            mdesc mMdesc
            num nActionIndex
            num nDelay = 0.5
            num nMoveType = 7
            num nPercentage
            num nSigValue
        pointRx pPointRx[2]
        string sID
      [5]
        bool bMarked
        jointRx jJointRx
        pointRx pInter
        paraItem pParaItem
          [0]
            bool bSafePoint
            ifItem iIfItem
              [0]
                bool bANDOR[2]
                num nSigIndex[3]
                num nSigType[3]
                num nValue[3]
            mdesc mMdesc
            num nActionIndex = 40
            num nDelay
            num nMoveType = 4
            num nPercentage
            num nSigValue
        pointRx pPointRx[2]
        string sID
    string sID
  [Y006]
    num nFrameIndex
    num nMoveID
    num nToolIndex
    pointItem pPointItem[6]
      [0]
        bool bMarked
        jointRx jJointRx
        pointRx pInter
        paraItem pParaItem
          [0]
            bool bSafePoint
            ifItem iIfItem
              [0]
                bool bANDOR[2]
                num nSigIndex[3]
                num nSigType[3]
                num nValue[3]
            mdesc mMdesc
            num nActionIndex = 40
            num nDelay
            num nMoveType = 4
            num nPercentage
            num nSigValue = 1
        pointRx pPointRx[2]
        string sID
      [1]
        bool bMarked
        jointRx jJointRx
        pointRx pInter
        paraItem pParaItem
          [0]
            bool bSafePoint
            ifItem iIfItem
              [0]
                bool bANDOR[2]
                num nSigIndex[3]
                num nSigType[3]
                num nValue[3]
            mdesc mMdesc
            num nActionIndex = 5
            num nDelay
            num nMoveType = 6
            num nPercentage
            num nSigValue = 6
        pointRx pPointRx[2]
        string sID
      [2]
        bool bMarked
        jointRx jJointRx
        pointRx pInter
        paraItem pParaItem
          [0]
            bool bSafePoint
            ifItem iIfItem
              [0]
                bool bANDOR[2]
                num nSigIndex[3]
                num nSigType[3]
                num nValue[3]
            mdesc mMdesc
            num nActionIndex
            num nDelay = 0.5
            num nMoveType = 7
            num nPercentage
            num nSigValue
        pointRx pPointRx[2]
        string sID
      [3]
        bool bMarked
        jointRx jJointRx
        pointRx pInter
        paraItem pParaItem
          [0]
            bool bSafePoint
            ifItem iIfItem
              [0]
                bool bANDOR[2]
                num nSigIndex[3]
                num nSigType[3]
                num nValue[3]
            mdesc mMdesc
            num nActionIndex = 40
            num nDelay = 0.5
            num nMoveType = 3
            num nPercentage
            num nSigValue = 1
        pointRx pPointRx[2]
        string sID
      [4]
        bool bMarked
        jointRx jJointRx
        pointRx pInter
        paraItem pParaItem
          [0]
            bool bSafePoint
            ifItem iIfItem
              [0]
                bool bANDOR[2]
                num nSigIndex[3]
                num nSigType[3]
                num nValue[3]
            mdesc mMdesc
            num nActionIndex
            num nDelay = 0.5
            num nMoveType = 7
            num nPercentage
            num nSigValue
        pointRx pPointRx[2]
        string sID
      [5]
        bool bMarked
        jointRx jJointRx
        pointRx pInter
        paraItem pParaItem
          [0]
            bool bSafePoint
            ifItem iIfItem
              [0]
                bool bANDOR[2]
                num nSigIndex[3]
                num nSigType[3]
                num nValue[3]
            mdesc mMdesc
            num nActionIndex = 40
            num nDelay
            num nMoveType = 4
            num nPercentage
            num nSigValue
        pointRx pPointRx[2]
        string sID
    string sID
  [Y007]
    num nFrameIndex
    num nMoveID
    num nToolIndex
    pointItem pPointItem[6]
      [0]
        bool bMarked
        jointRx jJointRx
        pointRx pInter
        paraItem pParaItem
          [0]
            bool bSafePoint
            ifItem iIfItem
              [0]
                bool bANDOR[2]
                num nSigIndex[3]
                num nSigType[3]
                num nValue[3]
            mdesc mMdesc
            num nActionIndex = 40
            num nDelay
            num nMoveType = 4
            num nPercentage
            num nSigValue = 1
        pointRx pPointRx[2]
        string sID
      [1]
        bool bMarked
        jointRx jJointRx
        pointRx pInter
        paraItem pParaItem
          [0]
            bool bSafePoint
            ifItem iIfItem
              [0]
                bool bANDOR[2]
                num nSigIndex[3]
                num nSigType[3]
                num nValue[3]
            mdesc mMdesc
            num nActionIndex = 5
            num nDelay
            num nMoveType = 6
            num nPercentage
            num nSigValue = 7
        pointRx pPointRx[2]
        string sID
      [2]
        bool bMarked
        jointRx jJointRx
        pointRx pInter
        paraItem pParaItem
          [0]
            bool bSafePoint
            ifItem iIfItem
              [0]
                bool bANDOR[2]
                num nSigIndex[3]
                num nSigType[3]
                num nValue[3]
            mdesc mMdesc
            num nActionIndex
            num nDelay = 0.5
            num nMoveType = 7
            num nPercentage
            num nSigValue
        pointRx pPointRx[2]
        string sID
      [3]
        bool bMarked
        jointRx jJointRx
        pointRx pInter
        paraItem pParaItem
          [0]
            bool bSafePoint
            ifItem iIfItem
              [0]
                bool bANDOR[2]
                num nSigIndex[3]
                num nSigType[3]
                num nValue[3]
            mdesc mMdesc
            num nActionIndex = 40
            num nDelay = 0.5
            num nMoveType = 3
            num nPercentage
            num nSigValue = 1
        pointRx pPointRx[2]
        string sID
      [4]
        bool bMarked
        jointRx jJointRx
        pointRx pInter
        paraItem pParaItem
          [0]
            bool bSafePoint
            ifItem iIfItem
              [0]
                bool bANDOR[2]
                num nSigIndex[3]
                num nSigType[3]
                num nValue[3]
            mdesc mMdesc
            num nActionIndex
            num nDelay = 0.5
            num nMoveType = 7
            num nPercentage
            num nSigValue
        pointRx pPointRx[2]
        string sID
      [5]
        bool bMarked
        jointRx jJointRx
        pointRx pInter
        paraItem pParaItem
          [0]
            bool bSafePoint
            ifItem iIfItem
              [0]
                bool bANDOR[2]
                num nSigIndex[3]
                num nSigType[3]
                num nValue[3]
            mdesc mMdesc
            num nActionIndex = 40
            num nDelay
            num nMoveType = 4
            num nPercentage
            num nSigValue
        pointRx pPointRx[2]
        string sID
    string sID
  [Y008]
    num nFrameIndex
    num nMoveID
    num nToolIndex
    pointItem pPointItem[6]
      [0]
        bool bMarked
        jointRx jJointRx
        pointRx pInter
        paraItem pParaItem
          [0]
            bool bSafePoint
            ifItem iIfItem
              [0]
                bool bANDOR[2]
                num nSigIndex[3]
                num nSigType[3]
                num nValue[3]
            mdesc mMdesc
            num nActionIndex = 40
            num nDelay
            num nMoveType = 4
            num nPercentage
            num nSigValue = 1
        pointRx pPointRx[2]
        string sID
      [1]
        bool bMarked
        jointRx jJointRx
        pointRx pInter
        paraItem pParaItem
          [0]
            bool bSafePoint
            ifItem iIfItem
              [0]
                bool bANDOR[2]
                num nSigIndex[3]
                num nSigType[3]
                num nValue[3]
            mdesc mMdesc
            num nActionIndex = 5
            num nDelay
            num nMoveType = 6
            num nPercentage
            num nSigValue = 8
        pointRx pPointRx[2]
        string sID
      [2]
        bool bMarked
        jointRx jJointRx
        pointRx pInter
        paraItem pParaItem
          [0]
            bool bSafePoint
            ifItem iIfItem
              [0]
                bool bANDOR[2]
                num nSigIndex[3]
                num nSigType[3]
                num nValue[3]
            mdesc mMdesc
            num nActionIndex
            num nDelay = 0.5
            num nMoveType = 7
            num nPercentage
            num nSigValue
        pointRx pPointRx[2]
        string sID
      [3]
        bool bMarked
        jointRx jJointRx
        pointRx pInter
        paraItem pParaItem
          [0]
            bool bSafePoint
            ifItem iIfItem
              [0]
                bool bANDOR[2]
                num nSigIndex[3]
                num nSigType[3]
                num nValue[3]
            mdesc mMdesc
            num nActionIndex = 40
            num nDelay = 0.5
            num nMoveType = 3
            num nPercentage
            num nSigValue = 1
        pointRx pPointRx[2]
        string sID
      [4]
        bool bMarked
        jointRx jJointRx
        pointRx pInter
        paraItem pParaItem
          [0]
            bool bSafePoint
            ifItem iIfItem
              [0]
                bool bANDOR[2]
                num nSigIndex[3]
                num nSigType[3]
                num nValue[3]
            mdesc mMdesc
            num nActionIndex
            num nDelay = 0.5
            num nMoveType = 7
            num nPercentage
            num nSigValue
        pointRx pPointRx[2]
        string sID
      [5]
        bool bMarked
        jointRx jJointRx
        pointRx pInter
        paraItem pParaItem
          [0]
            bool bSafePoint
            ifItem iIfItem
              [0]
                bool bANDOR[2]
                num nSigIndex[3]
                num nSigType[3]
                num nValue[3]
            mdesc mMdesc
            num nActionIndex = 40
            num nDelay
            num nMoveType = 4
            num nPercentage
            num nSigValue
        pointRx pPointRx[2]
        string sID
    string sID
  [complete]
    num nFrameIndex
    num nMoveID
    num nToolIndex
    pointItem pPointItem[3]
      [0]
        bool bMarked
        jointRx jJointRx
        pointRx pInter
        paraItem pParaItem
          [0]
            bool bSafePoint
            ifItem iIfItem
              [0]
                bool bANDOR[2]
                num nSigIndex[3]
                num nSigType[3]
                num nValue[3]
            mdesc mMdesc
            num nActionIndex = 50
            num nDelay
            num nMoveType = 4
            num nPercentage
            num nSigValue = 1
        pointRx pPointRx[2]
        string sID
      [1]
        bool bMarked
        jointRx jJointRx
        pointRx pInter
        paraItem pParaItem
          [0]
            bool bSafePoint
            ifItem iIfItem
              [0]
                bool bANDOR[2]
                num nSigIndex[3]
                num nSigType[3]
                num nValue[3]
            mdesc mMdesc
            num nActionIndex = 50
            num nDelay = 3
            num nMoveType = 7
            num nPercentage
            num nSigValue = 1
        pointRx pPointRx[2]
        string sID
      [2]
        bool bMarked
        jointRx jJointRx
        pointRx pInter
        paraItem pParaItem
          [0]
            bool bSafePoint
            ifItem iIfItem
              [0]
                bool bANDOR[2]
                num nSigIndex[3]
                num nSigType[3]
                num nValue[3]
            mdesc mMdesc
            num nActionIndex = 50
            num nDelay = 3
            num nMoveType = 4
            num nPercentage
            num nSigValue
        pointRx pPointRx[2]
        string sID
    string sID
  [gggg]
    num nFrameIndex
    num nMoveID
    num nToolIndex
    pointItem pPointItem
      [0]
        bool bMarked
        jointRx jJointRx
        pointRx pInter
        paraItem pParaItem
          [0]
            bool bSafePoint
            ifItem iIfItem
              [0]
                bool bANDOR[2]
                num nSigIndex[3]
                num nSigType[3]
                num nValue[3]
            mdesc mMdesc
            num nActionIndex
            num nDelay
            num nMoveType
            num nPercentage
            num nSigValue
        pointRx pPointRx[2]
        string sID
    string sID
  [init]
    num nFrameIndex
    num nMoveID
    num nToolIndex
    pointItem pPointItem[14]
      [0]
        bool bMarked
        jointRx jJointRx
        pointRx pInter
        paraItem pParaItem
          [0]
            bool bSafePoint
            ifItem iIfItem
              [0]
                bool bANDOR[2]
                num nSigIndex[3]
                num nSigType[3]
                num nValue[3]
            mdesc mMdesc
            num nActionIndex
            num nDelay
            num nMoveType = 6
            num nPercentage
            num nSigValue
        pointRx pPointRx[2]
        string sID
      [1]
        bool bMarked
        jointRx jJointRx
        pointRx pInter
        paraItem pParaItem
          [0]
            bool bSafePoint
            ifItem iIfItem
              [0]
                bool bANDOR[2]
                num nSigIndex[3]
                num nSigType[3]
                num nValue[3]
            mdesc mMdesc
            num nActionIndex = 3
            num nDelay
            num nMoveType = 6
            num nPercentage
            num nSigValue
        pointRx pPointRx[2]
        string sID
      [2]
        bool bMarked
        jointRx jJointRx
        pointRx pInter
        paraItem pParaItem
          [0]
            bool bSafePoint
            ifItem iIfItem
              [0]
                bool bANDOR[2]
                num nSigIndex[3]
                num nSigType[3]
                num nValue[3]
            mdesc mMdesc
            num nActionIndex = 2
            num nDelay
            num nMoveType = 6
            num nPercentage
            num nSigValue
        pointRx pPointRx[2]
        string sID
      [3]
        bool bMarked
        jointRx jJointRx
        pointRx pInter
        paraItem pParaItem
          [0]
            bool bSafePoint
            ifItem iIfItem
              [0]
                bool bANDOR[2]
                num nSigIndex[3]
                num nSigType[3]
                num nValue[3]
            mdesc mMdesc
            num nActionIndex = 1
            num nDelay
            num nMoveType = 6
            num nPercentage
            num nSigValue
        pointRx pPointRx[2]
        string sID
      [4]
        bool bMarked
        jointRx jJointRx
        pointRx pInter
        paraItem pParaItem
          [0]
            bool bSafePoint
            ifItem iIfItem
              [0]
                bool bANDOR[2]
                num nSigIndex[3]
                num nSigType[3]
                num nValue[3]
            mdesc mMdesc
            num nActionIndex = 4
            num nDelay
            num nMoveType = 6
            num nPercentage
            num nSigValue
        pointRx pPointRx[2]
        string sID
      [5]
        bool bMarked
        jointRx jJointRx
        pointRx pInter
        paraItem pParaItem
          [0]
            bool bSafePoint
            ifItem iIfItem
              [0]
                bool bANDOR[2]
                num nSigIndex[3]
                num nSigType[3]
                num nValue[3]
            mdesc mMdesc
            num nActionIndex = 5
            num nDelay
            num nMoveType = 6
            num nPercentage
            num nSigValue
        pointRx pPointRx[2]
        string sID
      [6]
        bool bMarked
        jointRx jJointRx
        pointRx pInter
        paraItem pParaItem
          [0]
            bool bSafePoint
            ifItem iIfItem
              [0]
                bool bANDOR[2]
                num nSigIndex[3]
                num nSigType[3]
                num nValue[3]
            mdesc mMdesc
            num nActionIndex = 50
            num nDelay
            num nMoveType = 4
            num nPercentage
            num nSigValue
        pointRx pPointRx[2]
        string sID
      [7]
        bool bMarked
        jointRx jJointRx
        pointRx pInter
        paraItem pParaItem
          [0]
            bool bSafePoint
            ifItem iIfItem
              [0]
                bool bANDOR[2]
                num nSigIndex[3]
                num nSigType[3]
                num nValue[3]
            mdesc mMdesc
            num nActionIndex = 40
            num nDelay
            num nMoveType = 4
            num nPercentage
            num nSigValue
        pointRx pPointRx[2]
        string sID
      [8]
        bool bMarked
        jointRx jJointRx
        pointRx pInter
        paraItem pParaItem
          [0]
            bool bSafePoint
            ifItem iIfItem
              [0]
                bool bANDOR[2]
                num nSigIndex[3]
                num nSigType[3]
                num nValue[3]
            mdesc mMdesc
            num nActionIndex = 41
            num nDelay
            num nMoveType = 4
            num nPercentage
            num nSigValue
        pointRx pPointRx[2]
        string sID
      [9]
        bool bMarked
        jointRx jJointRx
        pointRx pInter
        paraItem pParaItem
          [0]
            bool bSafePoint
            ifItem iIfItem
              [0]
                bool bANDOR[2]
                num nSigIndex[3]
                num nSigType[3]
                num nValue[3]
            mdesc mMdesc
            num nActionIndex = 42
            num nDelay
            num nMoveType = 4
            num nPercentage
            num nSigValue
        pointRx pPointRx[2]
        string sID
      [10]
        bool bMarked
        jointRx jJointRx
        pointRx pInter
        paraItem pParaItem
          [0]
            bool bSafePoint
            ifItem iIfItem
              [0]
                bool bANDOR[2]
                num nSigIndex[3]
                num nSigType[3]
                num nValue[3]
            mdesc mMdesc
            num nActionIndex = 43
            num nDelay
            num nMoveType = 4
            num nPercentage
            num nSigValue
        pointRx pPointRx[2]
        string sID
      [11]
        bool bMarked
        jointRx jJointRx
        pointRx pInter
        paraItem pParaItem
          [0]
            bool bSafePoint
            ifItem iIfItem
              [0]
                bool bANDOR[2]
                num nSigIndex[3]
                num nSigType[3]
                num nValue[3]
            mdesc mMdesc
            num nActionIndex = 44
            num nDelay
            num nMoveType = 4
            num nPercentage
            num nSigValue
        pointRx pPointRx[2]
        string sID
      [12]
        bool bMarked
        jointRx jJointRx
        pointRx pInter
        paraItem pParaItem
          [0]
            bool bSafePoint
            ifItem iIfItem
              [0]
                bool bANDOR[2]
                num nSigIndex[3]
                num nSigType[3]
                num nValue[3]
            mdesc mMdesc
            num nActionIndex = 47
            num nDelay
            num nMoveType = 4
            num nPercentage
            num nSigValue
        pointRx pPointRx[2]
        string sID
      [13]
        bool bMarked
        jointRx jJointRx
        pointRx pInter
        paraItem pParaItem
          [0]
            bool bSafePoint
            ifItem iIfItem
              [0]
                bool bANDOR[2]
                num nSigIndex[3]
                num nSigType[3]
                num nValue[3]
            mdesc mMdesc
            num nActionIndex = 48
            num nDelay
            num nMoveType = 4
            num nPercentage
            num nSigValue
        pointRx pPointRx[2]
        string sID
    string sID
  [p001]
    num nFrameIndex
    num nMoveID
    num nToolIndex
    pointItem pPointItem[109]
      [0]
        bool bMarked
        jointRx jJointRx = {j1=14.463054, j2=126.686617, j3=-94.408556, j4=-18.307578, j5=-113.737208, j6=85.971215}
        pointRx pInter
        paraItem pParaItem
          [0]
            bool bSafePoint
            ifItem iIfItem
              [0]
                bool bANDOR[2]
                num nSigIndex[3]
                num nSigType[3]
                num nValue[3]
            mdesc mMdesc
            num nActionIndex = 41
            num nDelay = 1
            num nMoveType = 7
            num nPercentage
            num nSigValue
        pointRx pPointRx[2] = {x=278.890712, y=136.745171, z=230.948915, rx=84.337923, ry=-1.664851, rz=172.690172, shoulder=lefty, elbow=enegative, wrist=wnegative}
        string sID
      [1]
        bool bMarked
        jointRx jJointRx = {j1=14.463054, j2=126.686617, j3=-94.408556, j4=-18.307578, j5=-113.737208, j6=85.971215}
        pointRx pInter
        paraItem pParaItem
          [0]
            bool bSafePoint
            ifItem iIfItem
              [0]
                bool bANDOR[2]
                num nSigIndex[3]
                num nSigType[3]
                num nValue[3]
            mdesc mMdesc
            num nActionIndex = 71
            num nDelay = 1
            num nMoveType = 4
            num nPercentage
            num nSigValue
        pointRx pPointRx[2] = {x=278.890712, y=136.745171, z=230.948915, rx=84.337923, ry=-1.664851, rz=172.690172, shoulder=lefty, elbow=enegative, wrist=wnegative}
        string sID
      [2]
        bool bMarked
        jointRx jJointRx = {j1=14.463054, j2=126.686617, j3=-94.408556, j4=-18.307578, j5=-113.737208, j6=85.971215}
        pointRx pInter
        paraItem pParaItem
          [0]
            bool bSafePoint
            ifItem iIfItem
              [0]
                bool bANDOR[2]
                num nSigIndex[3]
                num nSigType[3]
                num nValue[3]
            mdesc mMdesc
            num nActionIndex = 70
            num nDelay = 1
            num nMoveType = 4
            num nPercentage
            num nSigValue = 1
        pointRx pPointRx[2] = {x=278.890712, y=136.745171, z=230.948915, rx=84.337923, ry=-1.664851, rz=172.690172, shoulder=lefty, elbow=enegative, wrist=wnegative}
        string sID
      [3]
        bool bMarked
        jointRx jJointRx = {j1=14.463054, j2=126.686617, j3=-94.408556, j4=-18.307578, j5=-113.737208, j6=85.971215}
        pointRx pInter
        paraItem pParaItem
          [0]
            bool bSafePoint
            ifItem iIfItem
              [0]
                bool bANDOR[2]
                num nSigIndex[3]
                num nSigType[3]
                num nValue[3]
            mdesc mMdesc
            num nActionIndex = 70
            num nDelay = 1
            num nMoveType = 3
            num nPercentage
            num nSigValue = 1
        pointRx pPointRx[2] = {x=278.890712, y=136.745171, z=230.948915, rx=84.337923, ry=-1.664851, rz=172.690172, shoulder=lefty, elbow=enegative, wrist=wnegative}
        string sID
      [4]
        bool bMarked
        jointRx jJointRx = {j1=-0.746077, j2=38.654193, j3=103.0610419, j4=-179.633028, j5=123.454226, j6=8.386419}
        pointRx pInter
        paraItem pParaItem
          [0]
            bool bSafePoint
            ifItem iIfItem
              [0]
                bool bANDOR[2]
                num nSigIndex[3]
                num nSigType[3]
                num nValue[3]
            mdesc mMdesc = {leave=0}
            num nActionIndex = 41
            num nDelay = 1
            num nMoveType = 1
            num nPercentage
            num nSigValue
        pointRx pPointRx[2] = {x=872.305806, y=193.820048, z=536.464849, rx=0.56853, ry=18.254398, rz=-172.702509, shoulder=lefty, elbow=epositive, wrist=wpositive}
        string sID
      [5]
        bool bMarked
        jointRx jJointRx = {j1=51.683001, j2=14.0128577, j3=41.487368, j4=-190.116938, j5=47.437404, j6=-46.111455}
        pointRx pInter
        paraItem pParaItem
          [0]
            bool bSafePoint
            ifItem iIfItem
              [0]
                bool bANDOR[2]
                num nSigIndex[3]
                num nSigType[3]
                num nValue[3]
            mdesc mMdesc = {leave=0}
            num nActionIndex = 41
            num nDelay = 1
            num nMoveType = 1
            num nPercentage
            num nSigValue
        pointRx pPointRx[2] = {x=343.831478, y=794.97015, z=1353.817104, rx=-11.2659, ry=-0.603091, rz=179.184152, shoulder=lefty, elbow=epositive, wrist=wpositive}
        string sID
      [6]
        bool bMarked
        jointRx jJointRx = {j1=48.571653, j2=8.537471, j3=47.670319, j4=-192.590165, j5=47.244918, j6=-41.470425}
        pointRx pInter
        paraItem pParaItem
          [0]
            bool bSafePoint
            ifItem iIfItem
              [0]
                bool bANDOR[2]
                num nSigIndex[3]
                num nSigType[3]
                num nValue[3]
            mdesc mMdesc = {leave=0}
            num nActionIndex = 41
            num nDelay = 1
            num nMoveType = 1
            num nPercentage
            num nSigValue
        pointRx pPointRx[2] = {x=343.165039, y=762.685647, z=1347.441881, rx=-13.302409, ry=-0.597019, rz=179.189754, shoulder=lefty, elbow=epositive, wrist=wpositive}
        string sID
      [7]
        bool bMarked
        jointRx jJointRx = {j1=50.121421, j2=10.919611, j3=45.291003, j4=-186.538203, j5=51.209762, j6=-47.0163097}
        pointRx pInter
        paraItem pParaItem
          [0]
            bool bSafePoint
            ifItem iIfItem
              [0]
                bool bANDOR[2]
